                num nValue[3]
            mdesc mMdesc = {leave=0}
            num nActionIndex = 41
            num nDelay = 1
            num nMoveType = 1
            num nPercentage
            num nSigValue
        pointRx pPointRx[2] = {x=-80.977735, y=690.533781, z=996.975174, rx=-3.552851, ry=0.854955, rz=-0.845343, shoulder=lefty, elbow=epositive, wrist=wpositive}
        string sID
      [103]
        bool bMarked
        jointRx jJointRx = {j1=92.678654, j2=24.947285, j3=65.529789, j4=-178.978625, j5=86.968643, j6=86.426716}
        pointRx pInter
        paraItem pParaItem
          [0]
            bool bSafePoint
            ifItem iIfItem
              [0]
                bool bANDOR[2]
                num nSigIndex[3]
                num nSigType[3]
                num nValue[3]
            mdesc mMdesc = {leave=0}
            num nActionIndex = 41
            num nDelay = 1
            num nMoveType = 1
            num nPercentage
            num nSigValue
        pointRx pPointRx[2] = {x=-81.24855, y=685.152861, z=1057.497507, rx=-3.552668, ry=0.854951, rz=-0.845339, shoulder=lefty, elbow=epositive, wrist=wpositive}
        string sID
      [104]
        bool bMarked
        jointRx jJointRx = {j1=94.697022, j2=-26.101782, j3=117.801323, j4=-178.839759, j5=92.416802, j6=84.701619}
        pointRx pInter
        paraItem pParaItem
          [0]
            bool bSafePoint
            ifItem iIfItem
              [0]
                bool bANDOR[2]
                num nSigIndex[3]
                num nSigType[3]
                num nValue[3]
            mdesc mMdesc = {leave=0}
            num nActionIndex = 41
            num nDelay = 1
            num nMoveType = 1
            num nPercentage
            num nSigValue
        pointRx pPointRx[2] = {x=-70.0312042, y=207.928608, z=1030.831107, rx=0.620415, ry=1.214089, rz=-0.649604, shoulder=lefty, elbow=epositive, wrist=wpositive}
        string sID
      [105]
        bool bMarked
        jointRx jJointRx = {j1=-0.746077, j2=38.654194, j3=103.0610414, j4=-179.633029, j5=123.454226, j6=8.386419}
        pointRx pInter
        paraItem pParaItem
          [0]
            bool bSafePoint
            ifItem iIfItem
              [0]
                bool bANDOR[2]
                num nSigIndex[3]
                num nSigType[3]
                num nValue[3]
            mdesc mMdesc = {leave=0}
            num nActionIndex = 41
            num nDelay = 1
            num nMoveType = 1
            num nPercentage
            num nSigValue
        pointRx pPointRx[2] = {x=872.305806, y=193.820048, z=536.464849, rx=0.56853, ry=18.254398, rz=-172.702509, shoulder=lefty, elbow=epositive, wrist=wpositive}
        string sID
      [106]
        bool bMarked
        jointRx jJointRx = {j1=-0.746077, j2=38.654194, j3=103.0610414, j4=-179.633029, j5=123.454226, j6=8.386419}
        pointRx pInter
        paraItem pParaItem
          [0]
            bool bSafePoint
            ifItem iIfItem
              [0]
                bool bANDOR[2]
                num nSigIndex[3]
                num nSigType[3]
                num nValue[3]
            mdesc mMdesc = {leave=0}
            num nActionIndex = 71
            num nDelay = 1
            num nMoveType = 4
            num nPercentage
            num nSigValue
        pointRx pPointRx[2] = {x=872.305806, y=193.820048, z=536.464849, rx=0.56853, ry=18.254398, rz=-172.702509, shoulder=lefty, elbow=epositive, wrist=wpositive}
        string sID
      [107]
        bool bMarked
        jointRx jJointRx = {j1=-0.746077, j2=38.654194, j3=103.0610414, j4=-179.633029, j5=123.454226, j6=8.386419}
        pointRx pInter
        paraItem pParaItem
          [0]
            bool bSafePoint
            ifItem iIfItem
              [0]
                bool bANDOR[2]
                num nSigIndex[3]
                num nSigType[3]
                num nValue[3]
            mdesc mMdesc = {leave=0}
            num nActionIndex = 70
            num nDelay = 1
            num nMoveType = 4
            num nPercentage
            num nSigValue = 1
        pointRx pPointRx[2] = {x=872.305806, y=193.820048, z=536.464849, rx=0.56853, ry=18.254398, rz=-172.702509, shoulder=lefty, elbow=epositive, wrist=wpositive}
        string sID
      [108]
        bool bMarked
        jointRx jJointRx = {j1=-0.746077, j2=38.654194, j3=103.0610414, j4=-179.633029, j5=123.454226, j6=8.386419}
        pointRx pInter
        paraItem pParaItem
          [0]
            bool bSafePoint
            ifItem iIfItem
              [0]
                bool bANDOR[2]
                num nSigIndex[3]
                num nSigType[3]
                num nValue[3]
            mdesc mMdesc = {leave=0}
            num nActionIndex = 70
            num nDelay = 1
            num nMoveType = 3
            num nPercentage
            num nSigValue = 1
        pointRx pPointRx[2] = {x=872.305806, y=193.820048, z=536.464849, rx=0.56853, ry=18.254398, rz=-172.702509, shoulder=lefty, elbow=epositive, wrist=wpositive}
        string sID
    string sID
  [p002]
    num nFrameIndex
    num nMoveID
    num nToolIndex
    pointItem pPointItem[89]
      [0]
        bool bMarked
        jointRx jJointRx = {j1=1.472874, j2=128.415304, j3=-142.718421, j4=-10.676075, j5=-13.610921, j6=92.673149}
        pointRx pInter
        paraItem pParaItem
          [0]
            bool bSafePoint
            ifItem iIfItem
              [0]
                bool bANDOR[2]
                num nSigIndex[3]
                num nSigType[3]
                num nValue[3]
            mdesc mMdesc
            num nActionIndex = 60
            num nDelay = 1
            num nMoveType = 7
            num nPercentage
            num nSigValue = 1
        pointRx pPointRx[2] = {x=91.326194, y=-43.762939, z=599.882275, rx=-88.611323, ry=-173.490167, rz=-62.0834554, shoulder=lefty, elbow=enegative, wrist=wnegative}
        string sID
      [1]
        bool bMarked
        jointRx jJointRx = {j1=-0.746435, j2=38.656305, j3=103.0621354, j4=-179.633633, j5=123.453008, j6=8.386286}
        pointRx pInter
        paraItem pParaItem
          [0]
            bool bSafePoint
            ifItem iIfItem
              [0]
                bool bANDOR[2]
                num nSigIndex[3]
                num nSigType[3]
                num nValue[3]
            mdesc mMdesc = {leave=0}
            num nActionIndex = 60
            num nDelay = 1
            num nMoveType = 1
            num nPercentage
            num nSigValue = 1
        pointRx pPointRx[2] = {x=872.340958, y=193.819324, z=536.420305, rx=0.568193, ry=18.258826, rz=-172.70256, shoulder=lefty, elbow=epositive, wrist=wpositive}
        string sID
      [2]
        bool bMarked
        jointRx jJointRx = {j1=13.421878, j2=-4.818376, j3=127.477265, j4=-178.119237, j5=122.0948701, j6=-9.80116}
        pointRx pInter
        paraItem pParaItem
          [0]
            bool bSafePoint
            ifItem iIfItem
              [0]
                bool bANDOR[2]
                num nSigIndex[3]
                num nSigType[3]
                num nValue[3]
            mdesc mMdesc = {leave=0}
            num nActionIndex = 60
            num nDelay = 1
            num nMoveType = 1
            num nPercentage
            num nSigValue = 1
        pointRx pPointRx[2] = {x=448.783781, y=302.866041, z=805.255089, rx=1.42221, ry=0.904693, rz=-177.39771, shoulder=lefty, elbow=epositive, wrist=wpositive}
        string sID
      [3]
        bool bMarked
        jointRx jJointRx = {j1=-44.645904, j2=7.328511, j3=115.0443755, j4=-179.561776, j5=120.728528, j6=47.488337}
        pointRx pInter
        paraItem pParaItem
          [0]
            bool bSafePoint
            ifItem iIfItem
              [0]
                bool bANDOR[2]
                num nSigIndex[3]
                num nSigType[3]
                num nValue[3]
            mdesc mMdesc = {leave=0}
            num nActionIndex = 60
            num nDelay = 1
            num nMoveType = 1
            num nPercentage
            num nSigValue = 1
        pointRx pPointRx[2] = {x=448.783853, y=-225.927858, z=805.255091, rx=1.423155, ry=0.904518, rz=-177.398128, shoulder=lefty, elbow=epositive, wrist=wpositive}
        string sID
      [4]
        bool bMarked
        jointRx jJointRx = {j1=-62.817139, j2=-4.0550919, j3=114.877833, j4=-181.800671, j5=110.902525, j6=152.578279}
        pointRx pInter
        paraItem pParaItem
          [0]
            bool bSafePoint
            ifItem iIfItem
              [0]
                bool bANDOR[2]
                num nSigIndex[3]
                num nSigType[3]
                num nValue[3]
            mdesc mMdesc = {leave=0}
            num nActionIndex = 60
            num nDelay = 1
            num nMoveType = 1
            num nPercentage
            num nSigValue = 1
        pointRx pPointRx[2] = {x=141.309816, y=-439.69867, z=907.056828, rx=-0.847975, ry=1.455546, rz=-89.586771, shoulder=lefty, elbow=epositive, wrist=wpositive}
        string sID
      [5]
        bool bMarked
        jointRx jJointRx = {j1=-65.775154, j2=-11.286589, j3=121.17379, j4=-181.783018, j5=110.0548117, j6=155.568352}
        pointRx pInter
        paraItem pParaItem
          [0]
            bool bSafePoint
            ifItem iIfItem
              [0]
                bool bANDOR[2]
                num nSigIndex[3]
                num nSigType[3]
                num nValue[3]
            mdesc mMdesc = {leave=0}
            num nActionIndex = 60
            num nDelay = 1
            num nMoveType = 1
            num nPercentage
            num nSigValue = 1
        pointRx pPointRx[2] = {x=93.46676, y=-399.708918, z=907.0568192, rx=-0.848373, ry=1.454915, rz=-89.587006, shoulder=lefty, elbow=epositive, wrist=wpositive}
        string sID
      [6]
        bool bMarked
        jointRx jJointRx = {j1=-89.343726, j2=-14.0520862, j3=123.23006, j4=-181.559542, j5=110.00182126, j6=179.223519}
        pointRx pInter
        paraItem pParaItem
          [0]
            bool bSafePoint
            ifItem iIfItem
              [0]
                bool bANDOR[2]
                num nSigIndex[3]
                num nSigType[3]
                num nValue[3]
            mdesc mMdesc = {leave=0}
            num nActionIndex = 60
            num nDelay = 1
            num nMoveType = 1
            num nPercentage
            num nSigValue = 1
        pointRx pPointRx[2] = {x=-89.571375, y=-439.696116, z=908.183016, rx=-0.847403, ry=1.455842, rz=-89.586507, shoulder=lefty, elbow=epositive, wrist=wpositive}
        string sID
      [7]
        bool bMarked
        jointRx jJointRx = {j1=-97.996959, j2=-19.937374, j3=127.468112, j4=-181.395365, j5=108.567727, j6=187.966831}
        pointRx pInter
        paraItem pParaItem
          [0]
            bool bSafePoint
            ifItem iIfItem
              [0]
                bool bANDOR[2]
                num nSigIndex[3]
                num nSigType[3]
                num nValue[3]
            mdesc mMdesc = {leave=0}
            num nActionIndex = 60
            num nDelay = 1
            num nMoveType = 1
            num nPercentage
            num nSigValue = 1
        pointRx pPointRx[2] = {x=-151.396189, y=-399.203302, z=908.183017, rx=-0.847956, ry=1.454831, rz=-89.586993, shoulder=lefty, elbow=epositive, wrist=wpositive}
        string sID
      [8]
        bool bMarked
        jointRx jJointRx = {j1=-114.27656, j2=-17.103316, j3=125.494276, j4=-181.0386567, j5=109.759295, j6=204.339244}
        pointRx pInter
        paraItem pParaItem
          [0]
            bool bSafePoint
            ifItem iIfItem
              [0]
                bool bANDOR[2]
                num nSigIndex[3]
                num nSigType[3]
                num nValue[3]
            mdesc mMdesc = {leave=0}
            num nActionIndex = 60
            num nDelay = 1
            num nMoveType = 1
            num nPercentage
            num nSigValue = 1
        pointRx pPointRx[2] = {x=-273.810345, y=-400.0623046, z=908.183017, rx=-0.848201, ry=1.454846, rz=-89.587073, shoulder=lefty, elbow=epositive, wrist=wpositive}
        string sID
      [9]
        bool bMarked
        jointRx jJointRx = {j1=-127.657278, j2=-10.433545, j3=120.35131, j4=-180.680851, j5=111.476535, j6=217.81872}
        pointRx pInter
        paraItem pParaItem
          [0]
            bool bSafePoint
            ifItem iIfItem
              [0]
                bool bANDOR[2]
                num nSigIndex[3]
                num nSigType[3]
                num nValue[3]
            mdesc mMdesc = {leave=0}
            num nActionIndex = 60
            num nDelay = 1
            num nMoveType = 1
            num nPercentage
            num nSigValue = 1
        pointRx pPointRx[2] = {x=-396.27202, y=-400.0380268, z=908.183017, rx=-0.848146, ry=1.454711, rz=-89.587133, shoulder=lefty, elbow=epositive, wrist=wpositive}
        string sID
      [10]
        bool bMarked
        jointRx jJointRx = {j1=-128.36271, j2=-3.761737, j3=114.478235, j4=-180.664263, j5=112.282673, j6=218.521551}
        pointRx pInter
        paraItem pParaItem
          [0]
            bool bSafePoint
            ifItem iIfItem
              [0]
                bool bANDOR[2]
                num nSigIndex[3]
                num nSigType[3]
                num nValue[3]
            mdesc mMdesc = {leave=0}
            num nActionIndex = 60
            num nDelay = 1
            num nMoveType = 1
            num nPercentage
            num nSigValue = 1
        pointRx pPointRx[2] = {x=-435.458865, y=-440.104527, z=908.183014, rx=-0.847701, ry=1.454786, rz=-89.586922, shoulder=lefty, elbow=epositive, wrist=wpositive}
        string sID
      [11]
        bool bMarked
        jointRx jJointRx = {j1=-150.0477665, j2=-32.514416, j3=134.825133, j4=-179.992645, j5=103.995071, j6=240.452121}
        pointRx pInter
        paraItem pParaItem
          [0]
            bool bSafePoint
            ifItem iIfItem
              [0]
                bool bANDOR[2]
                num nSigIndex[3]
                num nSigType[3]
                num nValue[3]
            mdesc mMdesc = {leave=0}
            num nActionIndex = 60
            num nDelay = 1
            num nMoveType = 1
            num nPercentage
            num nSigValue = 1
        pointRx pPointRx[2] = {x=-395.783095, y=-194.614951, z=908.183017, rx=-0.847327, ry=1.455777, rz=-89.586554, shoulder=lefty, elbow=epositive, wrist=wpositive}
        string sID
      [12]
        bool bMarked
        jointRx jJointRx = {j1=-134.69585, j2=-46.818065, j3=140.758548, j4=-180.440291, j5=95.566393, j6=225.0617106}
        pointRx pInter
        paraItem pParaItem
          [0]
            bool bSafePoint
            ifItem iIfItem
              [0]
                bool bANDOR[2]
                num nSigIndex[3]
                num nSigType[3]
                num nValue[3]
            mdesc mMdesc = {leave=0}
            num nActionIndex = 60
            num nDelay = 1
            num nMoveType = 1
            num nPercentage
            num nSigValue = 1
        pointRx pPointRx[2] = {x=-273.822937, y=-193.801075, z=908.183004, rx=-0.847798, ry=1.45516, rz=-89.586883, shoulder=lefty, elbow=epositive, wrist=wpositive}
        string sID
      [13]
        bool bMarked
        jointRx jJointRx = {j1=-127.583198, j2=-59.931416, j3=144.313107, j4=-180.637226, j5=85.941253, j6=218.0391471}
        pointRx pInter
        paraItem pParaItem
          [0]
            bool bSafePoint
            ifItem iIfItem
              [0]
                bool bANDOR[2]
                num nSigIndex[3]
                num nSigType[3]
                num nValue[3]
            mdesc mMdesc = {leave=0}
            num nActionIndex = 60
            num nDelay = 1
            num nMoveType = 1
            num nPercentage
            num nSigValue = 1
        pointRx pPointRx[2] = {x=-205.507537, y=-153.186144, z=908.183015, rx=-0.848113, ry=1.45473, rz=-89.587038, shoulder=lefty, elbow=epositive, wrist=wpositive}
        string sID
      [14]
        bool bMarked
        jointRx jJointRx = {j1=-106.245156, j2=-54.130159, j3=142.943602, j4=-181.160225, j5=90.03352, j6=196.659426}
        pointRx pInter
        paraItem pParaItem
          [0]
            bool bSafePoint
            ifItem iIfItem
              [0]
                bool bANDOR[2]
                num nSigIndex[3]
                num nSigType[3]
                num nValue[3]
            mdesc mMdesc = {leave=0}
            num nActionIndex = 60
            num nDelay = 1
            num nMoveType = 1
            num nPercentage
            num nSigValue = 1
        pointRx pPointRx[2] = {x=-151.172217, y=-193.150052, z=908.183009, rx=-0.846797, ry=1.455202, rz=-89.586651, shoulder=lefty, elbow=epositive, wrist=wpositive}
        string sID
      [15]
        bool bMarked
        jointRx jJointRx = {j1=-88.181189, j2=-60.305543, j3=144.390904, j4=-181.487087, j5=84.888565, j6=178.726344}
        pointRx pInter
        paraItem pParaItem
          [0]
            bool bSafePoint
            ifItem iIfItem
              [0]
                bool bANDOR[2]
                num nSigIndex[3]
                num nSigType[3]
                num nValue[3]
            mdesc mMdesc = {leave=0}
            num nActionIndex = 60
            num nDelay = 1
            num nMoveType = 1
            num nPercentage
            num nSigValue = 1
        pointRx pPointRx[2] = {x=-89.569536, y=-153.278481, z=908.183005, rx=-0.848103, ry=1.454988, rz=-89.586955, shoulder=lefty, elbow=epositive, wrist=wpositive}
        string sID
      [16]
        bool bMarked
        jointRx jJointRx = {j1=-49.557544, j2=-34.484563, j3=135.784981, j4=-181.687213, j5=100.997091, j6=139.633512}
        pointRx pInter
        paraItem pParaItem
          [0]
            bool bSafePoint
            ifItem iIfItem
              [0]
                bool bANDOR[2]
                num nSigIndex[3]
                num nSigType[3]
                num nValue[3]
            mdesc mMdesc = {leave=0}
            num nActionIndex = 60
            num nDelay = 1
            num nMoveType = 1
            num nPercentage
            num nSigValue = 1
        pointRx pPointRx[2] = {x=91.99085, y=-192.859385, z=908.183008, rx=-0.847307, ry=1.454124, rz=-89.587021, shoulder=lefty, elbow=epositive, wrist=wpositive}
        string sID
      [17]
        bool bMarked
        jointRx jJointRx = {j1=-38.259075, j2=-31.636106, j3=134.381133, j4=-181.602569, j5=102.121996, j6=128.316422}
        pointRx pInter
        paraItem pParaItem
          [0]
            bool bSafePoint
            ifItem iIfItem
              [0]
                bool bANDOR[2]
                num nSigIndex[3]
                num nSigType[3]
                num nValue[3]
            mdesc mMdesc = {leave=0}
            num nActionIndex = 60
            num nDelay = 1
            num nMoveType = 1
            num nPercentage
            num nSigValue = 1
        pointRx pPointRx[2] = {x=140.816821, y=-153.701987, z=908.183017, rx=-0.847662, ry=1.455654, rz=-89.586815, shoulder=lefty, elbow=epositive, wrist=wpositive}
        string sID
      [18]
        bool bMarked
        jointRx jJointRx = {j1=-40.179142, j2=-27.276637, j3=132.0274318, j4=-181.635185, j5=104.179865, j6=130.172936}
        pointRx pInter
        paraItem pParaItem
          [0]
            bool bSafePoint
            ifItem iIfItem
              [0]
                bool bANDOR[2]
                num nSigIndex[3]
                num nSigType[3]
                num nValue[3]
            mdesc mMdesc = {leave=0}
            num nActionIndex = 60
            num nDelay = 1
            num nMoveType = 1
            num nPercentage
            num nSigValue = 1
        pointRx pPointRx[2] = {x=157.0426787, y=-181.601488, z=908.183016, rx=-0.846776, ry=1.454662, rz=-89.586965, shoulder=lefty, elbow=epositive, wrist=wpositive}
        string sID
      [19]
        bool bMarked
        jointRx jJointRx = {j1=-35.580444, j2=-19.513295, j3=127.180796, j4=-181.605937, j5=106.969996, j6=125.504771}
        pointRx pInter
        paraItem pParaItem
          [0]
            bool bSafePoint
            ifItem iIfItem
              [0]
                bool bANDOR[2]
                num nSigIndex[3]
                num nSigType[3]
                num nValue[3]
            mdesc mMdesc = {leave=0}
            num nActionIndex = 60
            num nDelay = 1
            num nMoveType = 1
            num nPercentage
            num nSigValue = 1
        pointRx pPointRx[2] = {x=215.440719, y=-188.396141, z=908.183012, rx=-0.847349, ry=1.455713, rz=-89.586804, shoulder=lefty, elbow=epositive, wrist=wpositive}
        string sID
      [20]
        bool bMarked
        jointRx jJointRx = {j1=-46.861333, j2=-13.357926, j3=110.998877, j4=-181.655797, j5=97.261814, j6=137.0488022}
        pointRx pInter
        paraItem pParaItem
          [0]
            bool bSafePoint
            ifItem iIfItem
              [0]
                bool bANDOR[2]
                num nSigIndex[3]
                num nSigType[3]
                num nValue[3]
            mdesc mMdesc = {leave=0}
            num nActionIndex = 60
            num nDelay = 1
            num nMoveType = 1
            num nPercentage
            num nSigValue = 1
        pointRx pPointRx[2] = {x=219.716515, y=-307.982599, z=1017.163748, rx=-0.848894, ry=1.455617, rz=-89.586999, shoulder=lefty, elbow=epositive, wrist=wpositive}
        string sID
      [21]
        bool bMarked
        jointRx jJointRx = {j1=-50.556699, j2=-9.360644, j3=107.724248, j4=-181.67957, j5=98.0900481, j6=140.718516}
        pointRx pInter
        paraItem pParaItem
          [0]
            bool bSafePoint
            ifItem iIfItem
              [0]
                bool bANDOR[2]
                num nSigIndex[3]
                num nSigType[3]
                num nValue[3]
            mdesc mMdesc = {leave=0}
            num nActionIndex = 60
            num nDelay = 1
            num nMoveType = 1
            num nPercentage
            num nSigValue = 1
        pointRx pPointRx[2] = {x=219.716543, y=-356.481532, z=1017.163754, rx=-0.848073, ry=1.45566, rz=-89.587058, shoulder=lefty, elbow=epositive, wrist=wpositive}
        string sID
      [22]
        bool bMarked
        jointRx jJointRx = {j1=-63.140376, j2=-19.0449446, j3=115.233116, j4=-181.690981, j5=96.284673, j6=153.358529}
        pointRx pInter
        paraItem pParaItem
          [0]
            bool bSafePoint
            ifItem iIfItem
              [0]
                bool bANDOR[2]
                num nSigIndex[3]
                num nSigType[3]
                num nValue[3]
            mdesc mMdesc = {leave=0}
            num nActionIndex = 60
            num nDelay = 1
            num nMoveType = 1
            num nPercentage
            num nSigValue = 1
        pointRx pPointRx[2] = {x=95.813985, y=-356.481498, z=1017.163748, rx=-0.848073, ry=1.454616, rz=-89.587374, shoulder=lefty, elbow=epositive, wrist=wpositive}
        string sID
      [23]
        bool bMarked
        jointRx jJointRx = {j1=-79.728318, j2=-26.048727, j3=119.787691, j4=-181.587117, j5=94.312383, j6=170.0187689}
        pointRx pInter
        paraItem pParaItem
          [0]
            bool bSafePoint
            ifItem iIfItem
              [0]
                bool bANDOR[2]
                num nSigIndex[3]
                num nSigType[3]
                num nValue[3]
            mdesc mMdesc = {leave=0}
            num nActionIndex = 60
            num nDelay = 1
            num nMoveType = 1
            num nPercentage
            num nSigValue = 1
        pointRx pPointRx[2] = {x=-27.885141, y=-356.481499, z=1017.163752, rx=-0.848101, ry=1.454714, rz=-89.587352, shoulder=lefty, elbow=epositive, wrist=wpositive}
        string sID
      [24]
        bool bMarked
        jointRx jJointRx = {j1=-98.538538, j2=-28.494425, j3=121.213081, j4=-181.31556, j5=93.772464, j6=188.865913}
        pointRx pInter
        paraItem pParaItem
          [0]
            bool bSafePoint
            ifItem iIfItem
              [0]
                bool bANDOR[2]
                num nSigIndex[3]
                num nSigType[3]
                num nValue[3]
            mdesc mMdesc = {leave=0}
            num nActionIndex = 60
            num nDelay = 1
            num nMoveType = 1
            num nPercentage
            num nSigValue = 1
        pointRx pPointRx[2] = {x=-148.842085, y=-356.481513, z=1017.163754, rx=-0.848192, ry=1.454763, rz=-89.587369, shoulder=lefty, elbow=epositive, wrist=wpositive}
        string sID
      [25]
        bool bMarked
        jointRx jJointRx = {j1=-116.525543, j2=-25.666163, j3=119.557118, j4=-180.926658, j5=95.298865, j6=206.853059}
        pointRx pInter
        paraItem pParaItem
          [0]
            bool bSafePoint
            ifItem iIfItem
              [0]
                bool bANDOR[2]
                num nSigIndex[3]
                num nSigType[3]
                num nValue[3]
            mdesc mMdesc = {leave=0}
            num nActionIndex = 60
            num nDelay = 1
            num nMoveType = 1
            num nPercentage
            num nSigValue = 1
        pointRx pPointRx[2] = {x=-270.651747, y=-356.48152, z=1017.16375, rx=-0.848282, ry=1.454622, rz=-89.587473, shoulder=lefty, elbow=epositive, wrist=wpositive}
        string sID
      [26]
        bool bMarked
        jointRx jJointRx = {j1=-130.862945, j2=-18.445899, j3=114.810144, j4=-180.550576, j5=97.957003, j6=221.196075}
        pointRx pInter
        paraItem pParaItem
          [0]
            bool bSafePoint
            ifItem iIfItem
              [0]
                bool bANDOR[2]
                num nSigIndex[3]
                num nSigType[3]
                num nValue[3]
            mdesc mMdesc = {leave=0}
            num nActionIndex = 60
            num nDelay = 1
            num nMoveType = 1
            num nPercentage
            num nSigValue = 1
        pointRx pPointRx[2] = {x=-393.726947, y=-356.481515, z=1017.163742, rx=-0.848193, ry=1.45465, rz=-89.587465, shoulder=lefty, elbow=epositive, wrist=wpositive}
        string sID
      [27]
        bool bMarked
        jointRx jJointRx = {j1=-140.91448, j2=-8.959057, j3=107.381228, j4=-180.2633, j5=100.0860396, j6=231.274084}
        pointRx pInter
        paraItem pParaItem
          [0]
            bool bSafePoint
            ifItem iIfItem
              [0]
                bool bANDOR[2]
                num nSigIndex[3]
                num nSigType[3]
                num nValue[3]
            mdesc mMdesc = {leave=0}
            num nActionIndex = 60
            num nDelay = 1
            num nMoveType = 1
            num nPercentage
            num nSigValue = 1
        pointRx pPointRx[2] = {x=-513.86612, y=-356.481511, z=1017.163748, rx=-0.848031, ry=1.454987, rz=-89.587282, shoulder=lefty, elbow=epositive, wrist=wpositive}
        string sID
      [28]
        bool bMarked
        jointRx jJointRx = {j1=-153.0418655, j2=-18.291818, j3=114.699918, j4=-179.903722, j5=98.0918043, j6=243.463229}
        pointRx pInter
        paraItem pParaItem
          [0]
            bool bSafePoint
            ifItem iIfItem
              [0]
                bool bANDOR[2]
                num nSigIndex[3]
                num nSigType[3]
                num nValue[3]
            mdesc mMdesc = {leave=0}
            num nActionIndex = 60
            num nDelay = 1
            num nMoveType = 1
            num nPercentage
            num nSigValue = 1
        pointRx pPointRx[2] = {x=-513.879461, y=-236.101565, z=1017.176534, rx=-0.848451, ry=1.457487, rz=-89.579995, shoulder=lefty, elbow=epositive, wrist=wpositive}
        string sID
      [29]
        bool bMarked
        jointRx jJointRx = {j1=-144.0175069, j2=-30.466025, j3=122.301625, j4=-180.170967, j5=93.514082, j6=234.419036}
        pointRx pInter
        paraItem pParaItem
          [0]
            bool bSafePoint
            ifItem iIfItem
              [0]
                bool bANDOR[2]
                num nSigIndex[3]
                num nSigType[3]
                num nValue[3]
            mdesc mMdesc = {leave=0}
            num nActionIndex = 60
            num nDelay = 1
            num nMoveType = 1
            num nPercentage
            num nSigValue = 1
        pointRx pPointRx[2] = {x=-395.442895, y=-236.101476, z=1017.176542, rx=-0.848256, ry=1.458452, rz=-89.579694, shoulder=lefty, elbow=epositive, wrist=wpositive}
        string sID
      [30]
        bool bMarked
        jointRx jJointRx = {j1=-128.64916, j2=-40.787631, j3=127.162043, j4=-180.609644, j5=87.947622, j6=219.0888357}
        pointRx pInter
        paraItem pParaItem
          [0]
            bool bSafePoint
            ifItem iIfItem
              [0]
                bool bANDOR[2]
                num nSigIndex[3]
                num nSigType[3]
                num nValue[3]
            mdesc mMdesc = {leave=0}
            num nActionIndex = 60
            num nDelay = 1
            num nMoveType = 1
            num nPercentage
            num nSigValue = 1
        pointRx pPointRx[2] = {x=-275.671993, y=-236.101428, z=1017.176549, rx=-0.848143, ry=1.458263, rz=-89.579729, shoulder=lefty, elbow=epositive, wrist=wpositive}
        string sID
      [31]
        bool bMarked
        jointRx jJointRx = {j1=-102.719844, j2=-45.653614, j3=128.986999, j4=-181.241518, j5=84.483238, j6=193.26102}
        pointRx pInter
        paraItem pParaItem
          [0]
            bool bSafePoint
            ifItem iIfItem
              [0]
                bool bANDOR[2]
                num nSigIndex[3]
                num nSigType[3]
                num nValue[3]
            mdesc mMdesc = {leave=0}
            num nActionIndex = 60
            num nDelay = 1
            num nMoveType = 1
            num nPercentage
            num nSigValue = 1
        pointRx pPointRx[2] = {x=-148.462899, y=-236.101436, z=1017.176557, rx=-0.848273, ry=1.458323, rz=-89.579789, shoulder=lefty, elbow=epositive, wrist=wpositive}
        string sID
      [32]
        bool bMarked
        jointRx jJointRx = {j1=-75.234087, j2=-41.778931, j3=127.557239, j4=-181.629427, j5=86.228668, j6=165.75692}
        pointRx pInter
        paraItem pParaItem
          [0]
            bool bSafePoint
            ifItem iIfItem
              [0]
                bool bANDOR[2]
                num nSigIndex[3]
                num nSigType[3]
                num nValue[3]
            mdesc mMdesc = {leave=0}
            num nActionIndex = 60
            num nDelay = 1
            num nMoveType = 1
            num nPercentage
            num nSigValue = 1
        pointRx pPointRx[2] = {x=-28.693584, y=-236.101465, z=1017.176551, rx=-0.84848, ry=1.457801, rz=-89.579944, shoulder=lefty, elbow=epositive, wrist=wpositive}
        string sID
      [33]
        bool bMarked
        jointRx jJointRx = {j1=-54.0547334, j2=-31.651411, j3=122.930841, j4=-181.679125, j5=91.109632, j6=144.429098}
        pointRx pInter
        paraItem pParaItem
          [0]
            bool bSafePoint
            ifItem iIfItem
              [0]
                bool bANDOR[2]
                num nSigIndex[3]
                num nSigType[3]
                num nValue[3]
            mdesc mMdesc = {leave=0}
            num nActionIndex = 60
            num nDelay = 1
            num nMoveType = 1
            num nPercentage
            num nSigValue = 1
        pointRx pPointRx[2] = {x=93.915656, y=-236.10152, z=1017.176542, rx=-0.848626, ry=1.458442, rz=-89.579827, shoulder=lefty, elbow=epositive, wrist=wpositive}
        string sID
      [34]
        bool bMarked
        jointRx jJointRx = {j1=-40.485912, j2=-18.976357, j3=115.184667, j4=-181.599954, j5=95.647484, j6=130.730056}
        pointRx pInter
        paraItem pParaItem
          [0]
            bool bSafePoint
            ifItem iIfItem
              [0]
                bool bANDOR[2]
                num nSigIndex[3]
                num nSigType[3]
                num nValue[3]
            mdesc mMdesc = {leave=0}
            num nActionIndex = 60
            num nDelay = 1
            num nMoveType = 1
            num nPercentage
            num nSigValue = 1
        pointRx pPointRx[2] = {x=218.0172115, y=-236.101515, z=1017.176533, rx=-0.848556, ry=1.458479, rz=-89.579805, shoulder=lefty, elbow=epositive, wrist=wpositive}
        string sID
      [35]
        bool bMarked
        jointRx jJointRx = {j1=-56.332421, j2=-2.00588257, j3=98.357776, j4=-191.102312, j5=109.350057, j6=144.0440218}
        pointRx pInter
        paraItem pParaItem
          [0]
            bool bSafePoint
            ifItem iIfItem
              [0]
                bool bANDOR[2]
                num nSigIndex[3]
                num nSigType[3]
                num nValue[3]
            mdesc mMdesc = {leave=0}
            num nActionIndex = 60
            num nDelay = 1
            num nMoveType = 1
            num nPercentage
            num nSigValue = 1
        pointRx pPointRx[2] = {x=217.982076, y=-280.4862, z=1017.176427, rx=-16.836049, ry=1.457605, rz=-89.579964, shoulder=lefty, elbow=epositive, wrist=wpositive}
        string sID
      [36]
        bool bMarked
        jointRx jJointRx = {j1=-57.0892302, j2=-1.130905, j3=95.0181686, j4=-191.116073, j5=107.536619, j6=145.199111}
        pointRx pInter
        paraItem pParaItem
          [0]
            bool bSafePoint
            ifItem iIfItem
              [0]
                bool bANDOR[2]
                num nSigIndex[3]
                num nSigType[3]
                num nValue[3]
            mdesc mMdesc = {leave=0}
            num nActionIndex = 60
            num nDelay = 1
            num nMoveType = 1
            num nPercentage
            num nSigValue = 1
        pointRx pPointRx[2] = {x=217.25826, y=-287.692057, z=1039.200253, rx=-17.404061, ry=1.458922, rz=-89.579582, shoulder=lefty, elbow=epositive, wrist=wpositive}
        string sID
      [37]
        bool bMarked
        jointRx jJointRx = {j1=-68.577465, j2=-8.930032, j3=102.19446, j4=-188.072592, j5=108.841438, j6=157.209783}
        pointRx pInter
        paraItem pParaItem
          [0]
            bool bSafePoint
            ifItem iIfItem
              [0]
                bool bANDOR[2]
                num nSigIndex[3]
                num nSigType[3]
                num nValue[3]
            mdesc mMdesc = {leave=0}
            num nActionIndex = 60
            num nDelay = 1
            num nMoveType = 1
            num nPercentage
            num nSigValue = 1
        pointRx pPointRx[2] = {x=92.341138, y=-287.692035, z=1039.200247, rx=-17.404564, ry=1.458107, rz=-89.579944, shoulder=lefty, elbow=epositive, wrist=wpositive}
        string sID
      [38]
        bool bMarked
        jointRx jJointRx = {j1=-82.103588, j2=-13.996174, j3=106.344491, j4=-184.0287877, j5=109.361575, j6=171.532972}
        pointRx pInter
        paraItem pParaItem
          [0]
            bool bSafePoint
            ifItem iIfItem
              [0]
                bool bANDOR[2]
                num nSigIndex[3]
                num nSigType[3]
                num nValue[3]
            mdesc mMdesc = {leave=0}
            num nActionIndex = 60
            num nDelay = 1
            num nMoveType = 1
            num nPercentage
            num nSigValue = 1
        pointRx pPointRx[2] = {x=-29.398116, y=-287.692032, z=1039.200246, rx=-17.40454, ry=1.458076, rz=-89.57997, shoulder=lefty, elbow=epositive, wrist=wpositive}
        string sID
      [39]
        bool bMarked
        jointRx jJointRx = {j1=-97.0207895, j2=-15.676372, j3=107.633001, j4=-179.313083, j5=109.407544, j6=187.346174}
        pointRx pInter
        paraItem pParaItem
          [0]
            bool bSafePoint
            ifItem iIfItem
              [0]
                bool bANDOR[2]
                num nSigIndex[3]
                num nSigType[3]
                num nValue[3]
            mdesc mMdesc = {leave=0}
            num nActionIndex = 60
            num nDelay = 1
            num nMoveType = 1
            num nPercentage
            num nSigValue = 1
        pointRx pPointRx[2] = {x=-151.844236, y=-287.692004, z=1039.200243, rx=-17.404828, ry=1.457352, rz=-89.580353, shoulder=lefty, elbow=epositive, wrist=wpositive}
        string sID
      [40]
        bool bMarked
        jointRx jJointRx = {j1=-111.45415, j2=-13.551235, j3=105.99558, j4=-174.795071, j5=109.149535, j6=202.636872}
        pointRx pInter
        paraItem pParaItem
          [0]
            bool bSafePoint
            ifItem iIfItem
              [0]
                bool bANDOR[2]
                num nSigIndex[3]
                num nSigType[3]
                num nValue[3]
            mdesc mMdesc = {leave=0}
            num nActionIndex = 60
            num nDelay = 1
            num nMoveType = 1
            num nPercentage
            num nSigValue = 1
        pointRx pPointRx[2] = {x=-274.56659, y=-287.692024, z=1039.200241, rx=-17.405138, ry=1.457536, rz=-89.580306, shoulder=lefty, elbow=epositive, wrist=wpositive}
        string sID
      [41]
        bool bMarked
        jointRx jJointRx = {j1=-123.657855, j2=-8.168773, j3=101.535959, j4=-171.227841, j5=108.575909, j6=215.54185}
        pointRx pInter
        paraItem pParaItem
          [0]
            bool bSafePoint
            ifItem iIfItem
              [0]
                bool bANDOR[2]
                num nSigIndex[3]
                num nSigType[3]
                num nValue[3]
            mdesc mMdesc = {leave=0}
            num nActionIndex = 60
            num nDelay = 1
            num nMoveType = 1
            num nPercentage
            num nSigValue = 1
        pointRx pPointRx[2] = {x=-395.706047, y=-287.692007, z=1039.200232, rx=-17.404604, ry=1.457158, rz=-89.580476, shoulder=lefty, elbow=epositive, wrist=wpositive}
        string sID
      [42]
        bool bMarked
        jointRx jJointRx = {j1=-133.481098, j2=-0.271586, j3=94.00243485, j4=-168.691358, j5=107.220034, j6=225.754693}
